{attribute 'hide_all_locals'}
FUNCTION_BLOCK SetMacro
VAR_INPUT
	Start 							: BOOL;
	OutputType 						: OUTPUT_ENUM;
	ActionType						: OUTPUT_ACTION_ENUM;
	TimeOutTime						: TIME;
	PostDelay						: TIME;
	FeedBack						: POINTER TO BOOL;
	SetOutput 						: POINTER TO BOOL;
	ResetOutput 					: POINTER TO BOOL;
END_VAR

VAR_OUTPUT
	Busy 							: BOOL;
	Done							: BOOL;
	Error 							: BOOL;
END_VAR
VAR
	state 							: UINT;
	fbStartTrigger					: R_TRIG;
	startTriggerOutput				: BOOL;
	fbTimerOn 						: TON;
	fbTimerOnStart					: BOOL;
	fbTimerOnEnd 					: BOOL;
	fbPostTimer						: TON;
	fbPostTimerOnStart				: BOOL;
	fbPostTimerOnEnd				: BOOL;
END_VAR

fbTimerOn(IN:=fbTimerOnStart, PT := TimeOutTime, Q => fbTimerOnEnd);
fbPostTimer(IN:=fbPostTimerOnStart, PT := PostDelay, Q => fbPostTimerOnEnd);
fbStartTrigger(CLK := Start, Q => startTriggerOutput);

CASE state OF
	(************************** state 0 - IDLE *************************)  
	0:	
		Busy := FALSE;
		Done := FALSE;
		Error := FALSE;
		
		IF startTriggerOutput THEN
			Busy := TRUE;
			Error := FALSE;
			fbTimerOnStart := FALSE;
			state := 10;
		END_IF
	10:
		IF FeedBack^ THEN
			IF PostDelay <> T#0MS THEN
				fbPostTimerOnStart := TRUE;
				state := 30;
			ELSE
				state := 100;
			END_IF
		ELSE
			fbTimerOnStart := TRUE;
			state := 20;
		END_IF
	
	(************** state 20 - Set Output and wait for feedback *************)  
	20:
		CASE ActionType OF
			OUTPUT_ACTION_ENUM.SET:
				SetOutput^ := TRUE;
				IF OutputType = OUTPUT_ENUM.BISTABLE THEN
					ResetOutput^ := FALSE;
				END_IF

			OUTPUT_ACTION_ENUM.RESET:
				SetOutput^ := FALSE;
				IF OutputType = OUTPUT_ENUM.BISTABLE THEN
					ResetOutput^ := TRUE;
				END_IF
		END_CASE
		
		// Il timeout prevale anche se il feedback arriva nella stessa scansione.
		IF fbTimerOnEnd THEN
			fbTimerOnStart := FALSE;
			SetOutput^ := FALSE;
			ResetOutput^ := FALSE;
			state := 200;
		ELSIF FeedBack^ THEN
			fbTimerOnStart := FALSE;
			//SetOutput^ := FALSE;
			//ResetOutput^ := FALSE;
			
			IF PostDelay <> T#0MS THEN
				fbPostTimerOnStart := TRUE;
				state := 30;
			ELSE
				state := 100;
			END_IF
		END_IF
		
	(************** state 30 - Wait Post Time Delay *************)  
	30:
		IF fbPostTimerOnEnd THEN
			fbPostTimerOnStart := FALSE;
			state := 100;
		END_IF
	
	(************** state 100 - End *************)  
	100:
		Done := TRUE;
		state := 0;
	
	(************** state 100 - Error *************)  
	200:
		state := 0;
		Error := TRUE;
		
END_CASE

END_FUNCTION_BLOCK

(* stored: Version 1.1.0.1, ProductVersion 3.1.4024.12
   POU SetMacro: Id {90e18c29-98d4-4a47-a59b-8a74665e8cc7}, SpecialFunc None *)
